TYPE SimulatorCommand :
STRUCT
	version : UDINT;
	cycle : UDINT;
	plcTimeInNs : ULINT;
	// The wheels' actual speed, from the NC axes. The simulator moves the robot with it.
	leftWheelVelocityInMPerS : LREAL;
	rightWheelVelocityInMPerS : LREAL;
	isLeftDriveEnabled : BOOL;
	isRightDriveEnabled : BOOL;
	isLidarPowered : BOOL;
	estimatedPose : Pose2D;
END_STRUCT
END_TYPE

(* stored: Version 1.1.0.1, ProductVersion 3.1.4026.12
   DUT SimulatorCommand: Id {ef5ef6ff-8903-5410-9bba-2c75dd95eb39} *)
